SUBAPPLICATION Uebung_158_AX (* Übung zu FsMkDir/FsMove/FsDelete: Ordner anlegen, umbenennen, kopieren, löschen *)
  (* Standard: 61499-2; Description: Copyright (c) 2026 Meisterschulen am Ostbahnhof This program and the accompanying materials are made available under the terms of the Eclipse Public License 2.0 which is available at https://www.eclipse.org/legal/epl-2.0/ SPDX-License-Identifier: EPL-2.0 *)
  (* Version 1.0, 2026-11-26, Franz Höpfinger, Meisterschulen am Ostbahnhof, initial API and implementation and/or initial documentation *)
  PACKAGE Uebungen;
  IMPORT Uebungen::const::Uebung_150_159::FileServer::FS_A;
  IMPORT Uebungen::const::Uebung_150_159::FileServer::FS_ADD;
  IMPORT Uebungen::const::Uebung_150_159::FileServer::FS_B;
  IMPORT Uebungen::const::Uebung_150_159::FileServer::FS_C;
  IMPORT Uebungen::const::Uebung_150_159::FileServer::FS_FLT;
  IMPORT Uebungen::const::Uebung_150_159::FileServer::FS_LOKAL;
  IMPORT Uebungen::const::Uebung_150_159::FileServer::FS_ORDNER;
  IMPORT isobus::pgn::ISOUSERHOME_e::network;
  IMPORT isobus::pgn::ISO_CAN_NODE::NODE1;
  IMPORT logiBUS::io::DI::logiBUS_DI::Input_I1;
  IMPORT logiBUS::io::DI::logiBUS_DI::Input_I2;
  IMPORT logiBUS::io::DI::logiBUS_DI_Events::BUTTON_SINGLE_CLICK;
  IMPORT logiBUS::io::DQ::logiBUS_DO::Output_Q1;
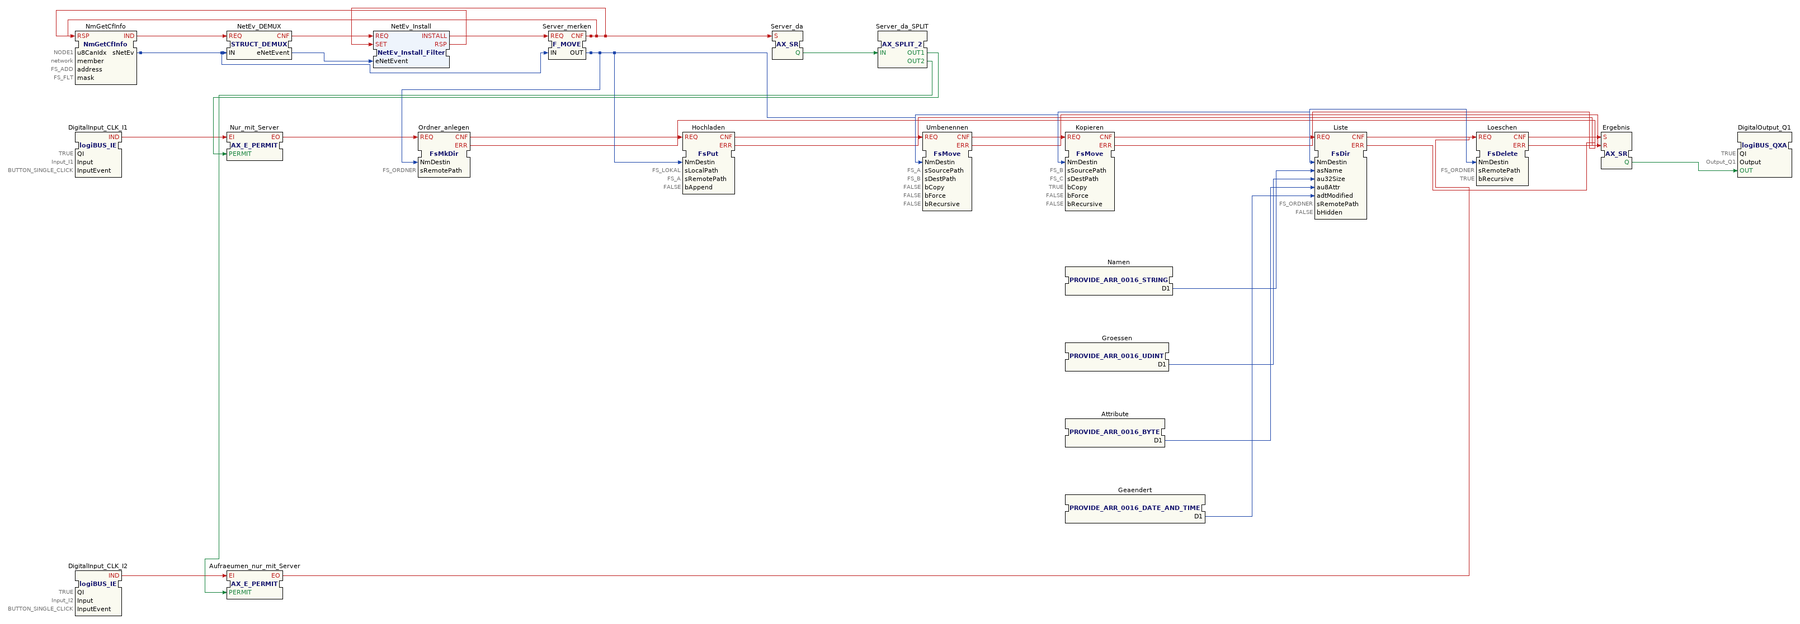
  (* File Server: Ordner anlegen, Datei umbenennen und kopieren, aufräumen (FsMkDir, FsPut, FsMove, FsDir, FsDelete) NmGetCfInfo (network, Filter FS_ADD/FS_FLT = NAME-Funktion 61) meldet den File Server, z. B. CCI 1200 mit USB-Stick. I1 Klick (nur mit Server): 1. FS_ORDNER anlegen, 2. FS_LOKAL nach a.txt, 3. a.txt in b.txt umbenennen, 4. b.txt nach c.txt kopieren, 5. Ordner listen, 6. Ordner löschen. Jeder Schritt startet nur nach CNF des vorigen. Bei ERR bleibt die Kette stehen: Q1 aus, s16Status und u16FsError des Schritts im Watch. I2 Klick: nur Ordner löschen. Offen am CCI 1200: Ordner anlegen (Schritt 1) und Kopieren (Schritt 4). FS_LOKAL muss es geben (Übung 156b). Voraussetzungen: Firmware mit den neuen File-Server-Bausteinen, neue isobus_fs-ELF, PART_13_FSC = 1 in /data/functionalities.ini. *)
  FBS
    NmGetCfInfo : isobus::pgn::NmGetCfInfo(u8CanIdx := NODE1, member := network, address := FS_ADD, mask := FS_FLT); (* meldet den File Server (Funktion 61) *)
    NetEv_DEMUX : eclipse4diac::convert::STRUCT_DEMUX; {SET_ATTRIBUTE(StructuredType, isobus::pgn::ISONETEVENT_T)}
    Server_merken : iec61131::selection::F_MOVE; (* eigener CF und File-Server-CF (NmDestin) *)
    Server_da : adapter::events::unidirectional::AX_SR;
    Server_da_SPLIT : adapter::events::unidirectional::AX_SPLIT_2;
    DigitalInput_CLK_I1 : logiBUS::io::DI::logiBUS_IE(QI := TRUE, Input := Input_I1, InputEvent := BUTTON_SINGLE_CLICK);
    Nur_mit_Server : adapter::events::unidirectional::AX_E_PERMIT;
    Ordner_anlegen : isobus::fs::FsMkDir(sRemotePath := FS_ORDNER); (* 1. FS_ORDNER anlegen *)
    Hochladen : isobus::fs::FsPut(sLocalPath := FS_LOKAL, sRemotePath := FS_A, bAppend := FALSE); (* 2. FS_LOKAL (aus Übung 156b) nach FS_A *)
    Umbenennen : isobus::fs::FsMove(sSourcePath := FS_A, sDestPath := FS_B, bCopy := FALSE, bForce := FALSE, bRecursive := FALSE); (* 3. FS_A in FS_B umbenennen *)
    Kopieren : isobus::fs::FsMove(sSourcePath := FS_B, sDestPath := FS_C, bCopy := TRUE, bForce := FALSE, bRecursive := FALSE); (* 4. FS_B nach FS_C kopieren (kann der CCI 1200 das?) *)
    Namen : eclipse4diac::convert::providers::PROVIDE_ARR_0016_STRING;
    Groessen : eclipse4diac::convert::providers::PROVIDE_ARR_0016_UDINT;
    Attribute : eclipse4diac::convert::providers::PROVIDE_ARR_0016_BYTE;
    Geaendert : eclipse4diac::convert::providers::PROVIDE_ARR_0016_DATE_AND_TIME;
    Liste : isobus::fs::FsDir(sRemotePath := FS_ORDNER, bHidden := FALSE); (* 5. FS_ORDNER listen (erwartet b.txt und c.txt) *)
    DigitalInput_CLK_I2 : logiBUS::io::DI::logiBUS_IE(QI := TRUE, Input := Input_I2, InputEvent := BUTTON_SINGLE_CLICK); (* nur Aufräumen, z. B. nach einem Fehler *)
    Aufraeumen_nur_mit_Server : adapter::events::unidirectional::AX_E_PERMIT;
    Loeschen : isobus::fs::FsDelete(sRemotePath := FS_ORDNER, bRecursive := TRUE); (* 6. FS_ORDNER mit Inhalt löschen *)
    Ergebnis : adapter::events::unidirectional::AX_SR; (* Q1 an = alle Schritte fertig *)
    DigitalOutput_Q1 : logiBUS::io::DQ::logiBUS_QXA(QI := TRUE, Output := Output_Q1);
  END_FBS
  SUBAPPS
    NetEv_Install : MyLib::sys::NetEv_Install_Filter;
  END_SUBAPPS
  EVENT_CONNECTIONS
    NmGetCfInfo.IND TO NetEv_DEMUX.REQ;
    NetEv_DEMUX.CNF TO NetEv_Install.REQ;
    NetEv_Install.INSTALL TO Server_merken.REQ;
    NetEv_Install.RSP TO NmGetCfInfo.RSP;
    Server_merken.CNF TO NetEv_Install.SET;
    Server_merken.CNF TO Server_da.S;
    Server_merken.CNF TO NmGetCfInfo.RSP;
    DigitalInput_CLK_I1.IND TO Nur_mit_Server.EI;
    Nur_mit_Server.EO TO Ordner_anlegen.REQ;
    Ordner_anlegen.CNF TO Hochladen.REQ;
    Hochladen.CNF TO Umbenennen.REQ;
    Umbenennen.CNF TO Kopieren.REQ;
    Kopieren.CNF TO Liste.REQ;
    Liste.CNF TO Loeschen.REQ;
    DigitalInput_CLK_I2.IND TO Aufraeumen_nur_mit_Server.EI;
    Aufraeumen_nur_mit_Server.EO TO Loeschen.REQ;
    Loeschen.CNF TO Ergebnis.S;
    Ordner_anlegen.ERR TO Ergebnis.R;
    Hochladen.ERR TO Ergebnis.R;
    Umbenennen.ERR TO Ergebnis.R;
    Kopieren.ERR TO Ergebnis.R;
    Liste.ERR TO Ergebnis.R;
    Loeschen.ERR TO Ergebnis.R;
  END_CONNECTIONS
  DATA_CONNECTIONS
    NmGetCfInfo.sNetEv TO NetEv_DEMUX.IN;
    NetEv_DEMUX.eNetEvent TO NetEv_Install.eNetEvent;
    NmGetCfInfo.sNetEv TO Server_merken.IN;
    Server_merken.OUT TO Ordner_anlegen.NmDestin;
    Server_merken.OUT TO Hochladen.NmDestin;
    Server_merken.OUT TO Umbenennen.NmDestin;
    Server_merken.OUT TO Kopieren.NmDestin;
    Server_merken.OUT TO Liste.NmDestin;
    Server_merken.OUT TO Loeschen.NmDestin;
    Namen.D1 TO Liste.asName;
    Groessen.D1 TO Liste.au32Size;
    Attribute.D1 TO Liste.au8Attr;
    Geaendert.D1 TO Liste.adtModified;
  END_CONNECTIONS
  ADAPTER_CONNECTIONS
    Server_da.Q TO Server_da_SPLIT.IN;
    Server_da_SPLIT.OUT1 TO Nur_mit_Server.PERMIT;
    Server_da_SPLIT.OUT2 TO Aufraeumen_nur_mit_Server.PERMIT;
    Ergebnis.Q TO DigitalOutput_Q1.OUT;
  END_CONNECTIONS
END_SUBAPPLICATION
